// TIA Portal V18 export
DATA_BLOCK "DB_MB_Comm_LoadConfig"   // DB5
{ S7_Optimized_Access := 'TRUE' }
// stored: MemoryReserve 0
   VAR
      BAUD : UDInt := 9600;
      PARITY : UInt;
      FLOW_CTRL : UInt;
      RTS_ON_DLY : UInt;
      RTS_OFF_DLY : UInt;
      RESP_TO : UInt := 1000;
      DONE : Bool;
      ERROR : Bool;
      STATUS : Word;
   END_VAR
BEGIN
END_DATA_BLOCK
